RoboDK station: PRBE_Tache_Bras.rdk

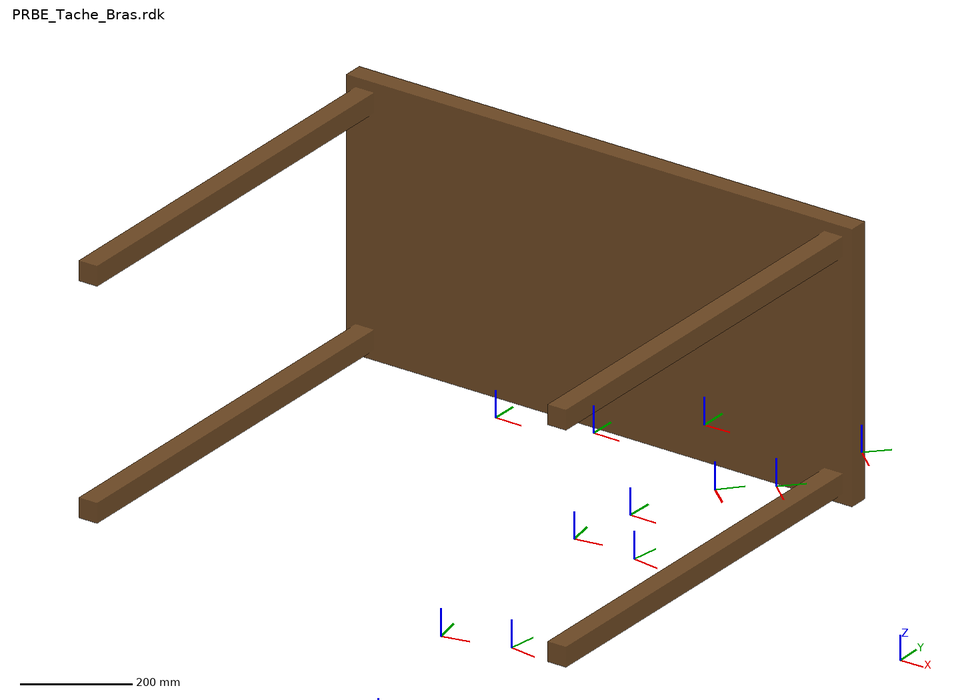
[picture v0: the station drawn from its stored meshes, robots at their saved joint values, targets as dots, program paths as lines]
Station PRBE_Tache_Bras (saved by RoboDK 6.0.4). Poses are relative to the parent item; angles as X-Y-Z fixed-axis rotations.
  - object Manikin_1 at (0, 0, 0) mm, geometry from Manikin_1.STEP
  - frame Human_Base at (0, 958, 0) mm
    - frame hipL_abduction at (63.26, -78.51, -37.42) mm, rotated rx 0 ry 0 rz -7.94 deg
      - frame hipL_flexion at (0, 0, 0) mm
        - frame hipL_rotation at (0, 0, 0) mm
          - frame kneeL_flexion at (67.44, -393.44, -12.97) mm
            - frame ankleL_flexion at (42.46, -394.54, 0) mm, rotated rx 0 ry 0 rz 7.94 deg
              - item type 7 Manikin_1-pied_g
            - item type 7 Manikin_1-tibia_g
          - item type 7 Manikin_1-cuisse_g
    - frame shoulderL_abduction at (206.4, 423.68, 12.96) mm, rotated rx 0 ry 0 rz -42 deg
      - frame shoulderL_flexion at (0, 0, 0) mm
        - frame shoulderL_rotation at (0, 0, 0) mm
          - frame elbowL_flexion at (155.8, -191.9, 27.9) mm
            - frame wristL_flexion at (148.7, -146.81, 80.89) mm
              - frame wristL_deviation at (0, 0, 0) mm
                - item type 7 Manikin_1-main_g
            - item type 7 Manikin_1-avant_bras_g
          - item type 7 Manikin_1-bras_g
    - frame hipR_abduction at (-70.11, -75.34, -37.06) mm, rotated rx 0 ry 0 rz 10.84 deg
      - frame hipR_flexion at (0, 0, 0) mm
        - frame hipR_rotation at (0, 0, 0) mm
          - frame kneeR_flexion at (-86.5, -385.51, -37.91) mm
            - frame ankleR_flexion at (-60.5, -382.31, -26.03) mm, rotated rx 0 ry 0 rz -10.84 deg
              - item type 7 Manikin_1-pied_d_1
              - item type 7 Manikin_1-pied_d_2
            - item type 7 Manikin_1-tibia_d_1
            - item type 7 Manikin_1-tibia_d_2
          - item type 7 Manikin_1-cuisse_d
    - frame shoulderR_abduction at (-133.98, 420.49, -26.02) mm
      - frame shoulderR_flexion at (0, 0, 0) mm
        - frame shoulderR_rotation at (0, 0, 0) mm
          - frame elbowR_flexion at (-80.76, -228.86, 52.14) mm
            - frame wristR_flexion at (-76.34, -195.54, 87.27) mm
              - frame wristR_deviation at (0, 0, 0) mm
                - item type 7 Manikin_1-main_d
            - item type 7 Manikin_1-avant_bras_d
          - item type 7 Manikin_1-bras_d
    - item type 7 Manikin_1-tete
    - item type 7 Manikin_1-bassin
    - item type 7 Manikin_1-torso
  - Python program Marche_Militaire (listed below)
  - Python program Marche_Avant (listed below)
  - Python program Marche_Trajectoire (listed below)
  - Python program fix_reattache_segments (listed below)
  - Python program Position_0 (listed below)
  - object Table at (0, 900, 485) mm, size 1100 x 900 x 550 mm
  - object Trajectoire_Marche at (0, 0, 0) mm
  - Python program Tache_Bras (listed below)
  - object Piece at (80, 940, 300) mm, size 80 x 80 x 80 mm

--- Python program Marche_Militaire ---
# -*- coding: utf-8 -*-
"""
Marche_Militaire.py — L'operateur marque le pas (marche militaire sur place).

A LANCER DANS ROBODK (clic droit > Run) depuis la station avec le rig 22 DDL,
operateur en pose NEUTRE (le script capture le repos au demarrage).

Principe de la marche militaire :
  - genoux qui montent haut, alternes
  - bras RAIDES (coude quasi tendu) qui balancent en OPPOSITION des jambes
  - buste droit (il est fige, parfait pour un militaire)

Regle les amplitudes/vitesse dans la section REGLAGES.
"""
from robolink import Robolink
from robodk.robomath import rotx, roty, rotz
import math
import time

RDK = Robolink()

# ---- Les 22 DDL : nom -> (axe, limite_basse_deg, limite_haute_deg) ----
DDL = {
    # JAMBE DROITE (5)
    "hipR_abduction": ("z", -45, 30),   "hipR_flexion": ("x", -120, 15),  "hipR_rotation": ("y", -45, 45),
    "kneeR_flexion":  ("x", 0, 135),    "ankleR_flexion": ("x", -30, 50),
    # JAMBE GAUCHE (5)
    "hipL_abduction": ("z", -30, 45),   "hipL_flexion": ("x", -120, 15),  "hipL_rotation": ("y", -45, 45),
    "kneeL_flexion":  ("x", 0, 135),    "ankleL_flexion": ("x", -30, 50),
    # BRAS DROIT (6)
    "shoulderR_abduction": ("z", -135, 90), "shoulderR_flexion": ("x", -90, 90), "shoulderR_rotation": ("y", -45, 180),
    "elbowR_flexion": ("x", 0, 145),
    "wristR_flexion": ("x", -50, 60),   "wristR_deviation": ("z", -30, 20),
    # BRAS GAUCHE (6)
    "shoulderL_abduction": ("z", -90, 135), "shoulderL_flexion": ("x", -90, 90), "shoulderL_rotation": ("y", -45, 180),
    "elbowL_flexion": ("x", 0, 145),
    "wristL_flexion": ("x", -50, 60),   "wristL_deviation": ("z", -30, 20),
}

ROT = {"x": rotx, "y": roty, "z": rotz}
F = {nom: RDK.Item(nom) for nom in DDL}            # les reperes
REST = {nom: F[nom].Pose() for nom in DDL}         # pose neutre (capturee au demarrage)


def bouge(nom, deg):
    """Tourne un DDL de `deg` degres depuis le repos (borne aux limites)."""
    axe, lo, hi = DDL[nom]
    deg = max(lo, min(hi, deg))
    F[nom].setPose(REST[nom] * ROT[axe](math.radians(deg)))


def neutre():
    """Remet tout l'operateur droit."""
    for nom in DDL:
        F[nom].setPose(REST[nom])


# =======================================================================
# REGLAGES de la marche militaire
# =======================================================================
HANCHE = 55      # levee de cuisse (deg) — genou haut
GENOU = 65       # pliage du genou quand la jambe monte (deg)
CHEVILLE = 15    # pointe de pied quand la jambe est levee (deg)
BRAS_AV = -45    # bras vers l'AVANT (deg, negatif = devant)
BRAS_ARR = 20    # bras vers l'ARRIERE (deg)
COUDE = 8        # coude quasi tendu = bras raide militaire
NB_PAS = 8       # nombre de pas au total
IMAGES_PAR_PAS = 12   # fluidite (images par pas)
DT = 0.04        # pause entre images (s) — plus petit = plus rapide


def pose_marche(ph):
    """Pose complete de la marche pour une phase `ph` (radians).
       Jambe droite levee sur [0, pi], jambe gauche sur [pi, 2pi]."""
    s = math.sin(ph)
    lift_d = max(0.0, s)     # jambe droite qui monte
    lift_g = max(0.0, -s)    # jambe gauche qui monte

    # jambes : genou haut + pointe de pied
    bouge("hipR_flexion", -HANCHE * lift_d)
    bouge("kneeR_flexion", GENOU * lift_d)
    bouge("ankleR_flexion", CHEVILLE * lift_d)
    bouge("hipL_flexion", -HANCHE * lift_g)
    bouge("kneeL_flexion", GENOU * lift_g)
    bouge("ankleL_flexion", CHEVILLE * lift_g)

    # bras raides, en opposition : bras droit devant quand jambe gauche monte
    u_d = (1.0 - s) / 2.0    # 0 = bras D derriere, 1 = bras D devant
    u_g = (1.0 + s) / 2.0
    bouge("shoulderR_flexion", BRAS_ARR + (BRAS_AV - BRAS_ARR) * u_d)
    bouge("shoulderL_flexion", BRAS_ARR + (BRAS_AV - BRAS_ARR) * u_g)
    bouge("elbowR_flexion", COUDE)
    bouge("elbowL_flexion", COUDE)


def marche(nb_pas=NB_PAS, images_par_pas=IMAGES_PAR_PAS, dt=DT):
    """Anime la marche militaire sur place."""
    for i in range(nb_pas * images_par_pas + 1):
        ph = math.pi * i / images_par_pas      # 1 pas = une demi-periode
        RDK.Render(False)
        pose_marche(ph)
        RDK.Render(True)
        time.sleep(dt)
    neutre()
    RDK.Render(True)


if __name__ == "__main__":
    print("Marche militaire : {} pas...".format(NB_PAS))
    marche()
    print("Repos !")

--- Python program Marche_Avant ---
# -*- coding: utf-8 -*-
"""
Marche_Avant.py — L'operateur marche TOUT DROIT devant lui (marche naturelle).

A LANCER DANS ROBODK (clic droit > Run) depuis la station avec le rig 22 DDL,
operateur au repos / garde-a-vous (le script capture le repos au demarrage).

Principe :
  - hanches qui balancent avant/arriere, genou qui se plie pendant le balance
  - bras souples en opposition des jambes (coude legerement plie)
  - le CORPS AVANCE a la vitesse des pas (longueur de pas calculee depuis
    l'amplitude de hanche) -> pas de glisse visible
  - il marche vers SON regard (+Z monde). A la fin, il REVIENT au centre
    (position d'origine de Human_Base).

Regle les amplitudes/vitesse dans la section REGLAGES.
"""
from robolink import Robolink
from robodk.robomath import rotx, roty, rotz, transl
import math
import time

RDK = Robolink()

# ---- Les 22 DDL : nom -> (axe, limite_basse_deg, limite_haute_deg) ----
DDL = {
    # JAMBE DROITE (5)
    "hipR_abduction": ("z", -45, 30),   "hipR_flexion": ("x", -120, 15),  "hipR_rotation": ("y", -45, 45),
    "kneeR_flexion":  ("x", 0, 135),    "ankleR_flexion": ("x", -30, 50),
    # JAMBE GAUCHE (5)
    "hipL_abduction": ("z", -30, 45),   "hipL_flexion": ("x", -120, 15),  "hipL_rotation": ("y", -45, 45),
    "kneeL_flexion":  ("x", 0, 135),    "ankleL_flexion": ("x", -30, 50),
    # BRAS DROIT (6)
    "shoulderR_abduction": ("z", -135, 90), "shoulderR_flexion": ("x", -90, 90), "shoulderR_rotation": ("y", -45, 180),
    "elbowR_flexion": ("x", 0, 145),
    "wristR_flexion": ("x", -50, 60),   "wristR_deviation": ("z", -30, 20),
    # BRAS GAUCHE (6)
    "shoulderL_abduction": ("z", -90, 135), "shoulderL_flexion": ("x", -90, 90), "shoulderL_rotation": ("y", -45, 180),
    "elbowL_flexion": ("x", 0, 145),
    "wristL_flexion": ("x", -50, 60),   "wristL_deviation": ("z", -30, 20),
}

ROT = {"x": rotx, "y": roty, "z": rotz}
F = {nom: RDK.Item(nom) for nom in DDL}            # les reperes
REST = {nom: F[nom].Pose() for nom in DDL}         # pose de repos (capturee au demarrage)
BASE = RDK.Item("Human_Base")
BASE_REST = BASE.Pose()                            # position de depart du corps
HOME = transl(0, 958, 0)                           # position d'origine (au centre, 1er repere)


def bouge(nom, deg):
    """Tourne un DDL de `deg` degres depuis le repos (borne aux limites)."""
    axe, lo, hi = DDL[nom]
    deg = max(lo, min(hi, deg))
    F[nom].setPose(REST[nom] * ROT[axe](math.radians(deg)))


def neutre():
    """Remet les articulations au repos (le corps reste ou il est)."""
    for nom in DDL:
        F[nom].setPose(REST[nom])


# =======================================================================
# REGLAGES de la marche
# =======================================================================
HANCHE_AV = 30    # jambe vers l'avant (deg)
HANCHE_ARR = 12   # jambe vers l'arriere (deg)
GENOU = 50        # pliage du genou pendant le balance (deg)
CHEVILLE = 8      # pointe de pied relevee pendant le balance (deg)
BRAS_AV = 25      # bras vers l'avant (deg)
BRAS_ARR = 15     # bras vers l'arriere (deg)
COUDE = 20        # coude legerement plie (marche naturelle)
NB_PAS = 8        # nombre de pas
IMAGES_PAR_PAS = 14   # fluidite
DT = 0.04         # pause entre images (s)

LONGUEUR_JAMBE = 790.0   # hanche -> cheville (mm, mesure sur le modele)
SENS = +1                # +1 = devant lui (+Z monde). Mets -1 pour marche arriere.

# longueur d'un pas deduite du balancement de hanche (pour avancer sans glisser)
LONGUEUR_PAS = LONGUEUR_JAMBE * (math.sin(math.radians(HANCHE_AV)) + math.sin(math.radians(HANCHE_ARR)))


def pose_pas(ph):
    """Pose de marche pour une phase `ph` (radians). Jambe droite devant sur [0, pi]."""
    s = math.sin(ph)
    # hanches : avant = negatif (amplitude asymetrique avant/arriere)
    a = (HANCHE_AV + HANCHE_ARR) / 2.0
    c = (HANCHE_AV - HANCHE_ARR) / 2.0
    bouge("hipR_flexion", -(a * s + c))
    bouge("hipL_flexion", -(a * -s + c))
    # genou plie pendant le balance (jambe qui revient vers l'avant)
    bouge("kneeR_flexion", GENOU * max(0.0, math.cos(ph)))
    bouge("kneeL_flexion", GENOU * max(0.0, -math.cos(ph)))
    # pointe de pied relevee pendant le balance (pour ne pas racler le sol)
    bouge("ankleR_flexion", -CHEVILLE * max(0.0, math.cos(ph)))
    bouge("ankleL_flexion", -CHEVILLE * max(0.0, -math.cos(ph)))
    # bras en opposition, coude souple
    sa = (BRAS_AV + BRAS_ARR) / 2.0
    sc = (BRAS_ARR - BRAS_AV) / 2.0
    bouge("shoulderR_flexion", sa * s + sc)
    bouge("shoulderL_flexion", -sa * s + sc)
    bouge("elbowR_flexion", COUDE)
    bouge("elbowL_flexion", COUDE)


def avance(dist):
    """Place le corps a `dist` mm devant sa position de depart."""
    BASE.setPose(BASE_REST * transl(0, 0, SENS * dist))


def marche(nb_pas=NB_PAS, images_par_pas=IMAGES_PAR_PAS, dt=DT):
    """Anime la marche en avant, puis remet l'operateur au centre (HOME)."""
    for i in range(nb_pas * images_par_pas + 1):
        ph = math.pi * i / images_par_pas      # 1 pas = une demi-periode
        RDK.Render(False)
        pose_pas(ph)
        avance(LONGUEUR_PAS * ph / math.pi)
        RDK.Render(True)
        time.sleep(dt)
    # fin : repos + retour a la position initiale, au centre
    RDK.Render(False)
    neutre()
    BASE.setPose(HOME)
    RDK.Render(True)


if __name__ == "__main__":
    d_tot = LONGUEUR_PAS * NB_PAS / 1000.0
    print("Marche avant : {} pas (~{:.1f} m)...".format(NB_PAS, d_tot))
    marche()
    print("Arrive !")

--- Python program Marche_Trajectoire ---
# -*- coding: utf-8 -*-
"""
Marche_Trajectoire.py — L'operateur marche le long d'une TRAJECTOIRE EXTERNE
(non lineaire), definie par des waypoints dans un fichier JSON.

A LANCER DANS ROBODK (clic droit > Run) depuis la station avec le rig 22 DDL,
operateur au repos / garde-a-vous (le script capture le repos au demarrage).

Principe (demande reunion du 04/06) :
  - la trajectoire est DEFINIE EN EXTERNE : trajectoires\\trajectoire_S.json
    (liste de points [x, z] au sol, en mm) -> modifiable sans toucher au code
  - les waypoints sont lisses par une spline Catmull-Rom -> courbe douce
  - le corps SUIT la courbe par abscisse curviligne : position sur la courbe
    + orientation vers la tangente (il regarde toujours ou il va)
  - meme cycle de marche et meme anti-glisse que Marche_Avant : le corps
    avance a la vitesse des pas (longueur de pas deduite du balancement
    de hanche), donc pas de patinage le long de la courbe
  - la trajectoire est tracee au sol dans la station (courbe bleue)

Usage terminal (RoboDK ouvert) :
    python Marche_Trajectoire.py [chemin\\trajectoire.json] [--reste]
    --reste : ne pas revenir au centre a la fin (rester au bout du chemin)
"""
from robolink import Robolink
from robodk.robomath import rotx, roty, rotz, transl
import bisect
import json
import math
import sys
import time

RDK = Robolink()

# ---- Les 22 DDL : nom -> (axe, limite_basse_deg, limite_haute_deg) ----
DDL = {
    # JAMBE DROITE (5)
    "hipR_abduction": ("z", -45, 30),   "hipR_flexion": ("x", -120, 15),  "hipR_rotation": ("y", -45, 45),
    "kneeR_flexion":  ("x", 0, 135),    "ankleR_flexion": ("x", -30, 50),
    # JAMBE GAUCHE (5)
    "hipL_abduction": ("z", -30, 45),   "hipL_flexion": ("x", -120, 15),  "hipL_rotation": ("y", -45, 45),
    "kneeL_flexion":  ("x", 0, 135),    "ankleL_flexion": ("x", -30, 50),
    # BRAS DROIT (6)
    "shoulderR_abduction": ("z", -135, 90), "shoulderR_flexion": ("x", -90, 90), "shoulderR_rotation": ("y", -45, 180),
    "elbowR_flexion": ("x", 0, 145),
    "wristR_flexion": ("x", -50, 60),   "wristR_deviation": ("z", -30, 20),
    # BRAS GAUCHE (6)
    "shoulderL_abduction": ("z", -90, 135), "shoulderL_flexion": ("x", -90, 90), "shoulderL_rotation": ("y", -45, 180),
    "elbowL_flexion": ("x", 0, 145),
    "wristL_flexion": ("x", -50, 60),   "wristL_deviation": ("z", -30, 20),
}

ROT = {"x": rotx, "y": roty, "z": rotz}
F = {nom: RDK.Item(nom) for nom in DDL}            # les reperes
REST = {nom: F[nom].Pose() for nom in DDL}         # pose de repos (capturee au demarrage)
BASE = RDK.Item("Human_Base")
HOME = transl(0, 958, 0)                           # position d'origine (au centre)
Y0 = BASE.Pose().Pos()[1]                          # hauteur du bassin (958 mm)


def bouge(nom, deg):
    """Tourne un DDL de `deg` degres depuis le repos (borne aux limites)."""
    axe, lo, hi = DDL[nom]
    deg = max(lo, min(hi, deg))
    F[nom].setPose(REST[nom] * ROT[axe](math.radians(deg)))


def neutre():
    """Remet les articulations au repos (le corps reste ou il est)."""
    for nom in DDL:
        F[nom].setPose(REST[nom])


# =======================================================================
# REGLAGES
# =======================================================================
TRAJET_DEFAUT = r"D:\PRBE_Homme_Robot\PRBE-Homme-Robot\trajectoires\trajectoire_S.json"
HANCHE_AV = 30    # jambe vers l'avant (deg)
HANCHE_ARR = 12   # jambe vers l'arriere (deg)
GENOU = 50        # pliage du genou pendant le balance (deg)
CHEVILLE = 8      # pointe de pied relevee pendant le balance (deg)
BRAS_AV = 25      # bras vers l'avant (deg)
BRAS_ARR = 15     # bras vers l'arriere (deg)
COUDE = 20        # coude legerement plie
IMAGES_PAR_PAS = 14   # fluidite
DT = 0.04         # pause entre images (s)
TRACER = True     # dessiner la trajectoire au sol dans la station

LONGUEUR_JAMBE = 790.0   # hanche -> cheville (mm)
LONGUEUR_PAS = LONGUEUR_JAMBE * (math.sin(math.radians(HANCHE_AV)) + math.sin(math.radians(HANCHE_ARR)))


# =======================================================================
# Trajectoire : JSON -> spline Catmull-Rom -> abscisse curviligne
# =======================================================================
def charge_waypoints(chemin):
    with open(chemin, encoding="utf-8") as f:
        data = json.load(f)
    pts = [tuple(map(float, p)) for p in data["points_xz_mm"]]
    if len(pts) < 2:
        raise SystemExit("ERREUR : il faut au moins 2 waypoints.")
    return data.get("nom", "(sans nom)"), pts


def _cr(p0, p1, p2, p3, t):
    """Point de Catmull-Rom (uniforme) entre p1 et p2, t dans [0,1]."""
    t2, t3 = t * t, t * t * t
    return tuple(0.5 * (2 * p1[k] + (-p0[k] + p2[k]) * t
                        + (2 * p0[k] - 5 * p1[k] + 4 * p2[k] - p3[k]) * t2
                        + (-p0[k] + 3 * p1[k] - 3 * p2[k] + p3[k]) * t3)
                 for k in range(2))


def lisse(waypoints, par_segment=24):
    """Spline Catmull-Rom a travers les waypoints -> polyligne dense."""
    P = [waypoints[0]] + list(waypoints) + [waypoints[-1]]
    dense = []
    for i in range(len(waypoints) - 1):
        for j in range(par_segment):
            dense.append(_cr(P[i], P[i + 1], P[i + 2], P[i + 3], j / par_segment))
    dense.append(waypoints[-1])
    return dense


def abscisses(dense):
    """Longueurs cumulees le long de la polyligne."""
    S = [0.0]
    for a, b in zip(dense, dense[1:]):
        S.append(S[-1] + math.hypot(b[0] - a[0], b[1] - a[1]))
    return S


def point_et_tangente(dense, S, s):
    """Position (x,z) + tangente unitaire (tx,tz) a l'abscisse s (mm)."""
    s = max(0.0, min(S[-1], s))
    i = min(max(bisect.bisect_left(S, s), 1), len(S) - 1)
    seg = S[i] - S[i - 1] or 1e-9
    u = (s - S[i - 1]) / seg
    a, b = dense[i - 1], dense[i]
    x = a[0] + u * (b[0] - a[0])
    z = a[1] + u * (b[1] - a[1])
    tx, tz = b[0] - a[0], b[1] - a[1]
    n = math.hypot(tx, tz) or 1e-9
    return (x, z), (tx / n, tz / n)


def tracer_trajectoire(dense):
    """Dessine la courbe au sol dans la station (best effort)."""
    try:
        vieux = RDK.Item("Trajectoire_Marche")
        if vieux.Valid() and vieux.Name() == "Trajectoire_Marche":
            vieux.Delete()
        courbe = RDK.AddCurve([[p[0], 10.0, p[1]] for p in dense])
        if courbe.Valid():
            courbe.setName("Trajectoire_Marche")
            courbe.setColorCurve([0.1, 0.3, 0.9, 1])
    except Exception as e:  # noqa: BLE001
        print("(trace de la trajectoire ignoree : {})".format(e))


# =======================================================================
# Cycle de marche (identique a Marche_Avant)
# =======================================================================
def pose_pas(ph):
    """Pose de marche pour une phase `ph` (radians). Jambe droite devant sur [0, pi]."""
    s = math.sin(ph)
    a = (HANCHE_AV + HANCHE_ARR) / 2.0
    c = (HANCHE_AV - HANCHE_ARR) / 2.0
    bouge("hipR_flexion", -(a * s + c))
    bouge("hipL_flexion", -(a * -s + c))
    bouge("kneeR_flexion", GENOU * max(0.0, math.cos(ph)))
    bouge("kneeL_flexion", GENOU * max(0.0, -math.cos(ph)))
    bouge("ankleR_flexion", -CHEVILLE * max(0.0, math.cos(ph)))
    bouge("ankleL_flexion", -CHEVILLE * max(0.0, -math.cos(ph)))
    sa = (BRAS_AV + BRAS_ARR) / 2.0
    sc = (BRAS_ARR - BRAS_AV) / 2.0
    bouge("shoulderR_flexion", sa * s + sc)
    bouge("shoulderL_flexion", -sa * s + sc)
    bouge("elbowR_flexion", COUDE)
    bouge("elbowL_flexion", COUDE)


def place_corps(dense, S, s):
    """Place le corps a l'abscisse s : position sur la courbe + regard tangent."""
    (x, z), (tx, tz) = point_et_tangente(dense, S, s)
    theta = math.atan2(tx, tz)          # le mannequin regarde vers +Z local
    BASE.setPose(transl(x, Y0, z) * roty(theta))


def marche_trajectoire(dense, S, retour_centre=True):
    """Anime la marche le long de la courbe, du debut a la fin."""
    L = S[-1]
    nb_images = int(math.ceil(L / LONGUEUR_PAS * IMAGES_PAR_PAS))
    for i in range(nb_images + 1):
        ph = math.pi * i / IMAGES_PAR_PAS          # 1 pas = une demi-periode
        s = min(L, LONGUEUR_PAS * ph / math.pi)    # anti-glisse : s = vitesse des pas
        RDK.Render(False)
        pose_pas(ph)
        place_corps(dense, S, s)
        RDK.Render(True)
        time.sleep(DT)
    # fin : repos (oriente comme a l'arrivee)
    RDK.Render(False)
    neutre()
    if retour_centre:
        BASE.setPose(HOME)
    RDK.Render(True)


if __name__ == "__main__":
    args = [a for a in sys.argv[1:] if a != "--reste"]
    reste = "--reste" in sys.argv[1:]
    chemin = args[0] if args else TRAJET_DEFAUT

    nom, waypoints = charge_waypoints(chemin)
    dense = lisse(waypoints)
    S = abscisses(dense)
    if TRACER:
        tracer_trajectoire(dense)
    print("Trajectoire '{}' : {} waypoints, {:.1f} m, ~{} pas".format(
        nom, len(waypoints), S[-1] / 1000.0, int(round(S[-1] / LONGUEUR_PAS))))
    marche_trajectoire(dense, S, retour_centre=not reste)
    p = BASE.Pose().Pos()
    print("Arrive ! Position finale Human_Base : x={:.0f} y={:.0f} z={:.0f} (retour_centre={})".format(
        p[0], p[1], p[2], not reste))

--- Python program fix_reattache_segments ---
# -*- coding: utf-8 -*-
"""
fix_reattache_segments.py — Repare le mannequin eclate a la reouverture du
.rdk SANS rebuild (quelques secondes), en re-jouant le re-basage geometrique
perdu a la sauvegarde.

Cause (diagnostic du 10/06) : pour les sous-solides type 7 (courbes issues
du Split), le .rdk sauve les points BRUTS d'origine — la compensation posee
par setParentStatic au moment du rig n'est PAS persistee. A l'ouverture,
RoboDK applique la transformation du frame parent sur ces points bruts
-> double transformation -> mannequin eclate. Les frames, vrais items a
pose persistee, restent corrects.

Remede, segment par segment :
  1) memoriser la pose relative de chaque frame, puis remettre chaque
     frame en etat de CONSTRUCTION (translation seule, rotation identite —
     l'etat dans lequel le rig d'origine a pose ses compensations)
  2) setParent(station)      — detache en KEEP-RELATIVE : la compensation
     (identite au chargement) ne change pas -> le segment retombe sur ses
     points bruts = position d'import, mannequin recompose
     setParentStatic(frame)  — re-attache en preservant l'absolu : la
     compensation F_build^-1 est re-posee, exactement comme au rig
  3) restaurer les poses memorisees (garde-a-vous, jambes resserrees) :
     la geometrie suit les frames

!! NE PAS envelopper dans RDK.Render(False) : le re-basage des type 7
echoue silencieusement sans rendu actif (constate le 10/06 — deux
tentatives identiques en Render(False) = aucun effet, la meme sequence
render actif fonctionne).

A relancer A CHAQUE OUVERTURE du .rdk (la sauvegarde re-perd le re-basage).
Filet de securite si etat incoherent : scripts/rebuild_operateur.py (~30 s).

!! PAS IDEMPOTENT : sur une station SAINE (fraichement rebuildee ou deja
reparee), le re-basage s'appliquerait une fois de trop et eclaterait le
mannequin. Une garde detecte l'etat via un segment du tronc et refuse de
tourner si la station est saine (--force pour outrepasser).

Usage (RoboDK ouvert, station chargee) :
    python fix_reattache_segments.py [--skip nom1,nom2] [--force]
    --skip  : segments a ne pas toucher (ex. deja repares a la main)
    --force : sauter la garde de detection
"""
import math
import sys
import time
from pathlib import Path
sys.path.insert(0, str(Path(__file__).resolve().parent))
from robolink import Robolink, ITEM_TYPE_FRAME
from robodk.robomath import transl

# ancres d'import des segments du tronc (cf. build_human_robodk.ANCHORS),
# en dur pour que le script reste autonome une fois embarque dans la station
TRONC = {"tete": (20, 1584, 30), "torso": (15, 1260, 0), "bassin": (0, 958, 0)}

skip = set()
if "--skip" in sys.argv:
    skip = set(sys.argv[sys.argv.index("--skip") + 1].split(","))

t0 = time.time()
RDK = Robolink()
station = RDK.ActiveStation()
print("Station :", station.Name())


def _d(a, b):
    return math.sqrt(sum((x - y) ** 2 for x, y in zip(a, b)))


def garde_station_cassee():
    """True si le mannequin est eclate (double transformation detectee)."""
    for it in RDK.ItemList():
        if it.Type() != 7:
            continue
        part = it.Name().split("-", 1)[-1]
        if part not in TRONC:
            continue
        bb = it.setParam("BoundingBox")
        c = [(bb["min"][i] + bb["max"][i]) / 2.0 for i in range(3)]
        a = TRONC[part]
        F = it.Parent().PoseAbs().rows
        fa = [sum(F[i][j] * a[j] for j in range(3)) + F[i][3] for i in range(3)]
        d_sain, d_casse = _d(c, a), _d(c, fa)
        etat = "CASSEE (double transformation)" if d_casse < d_sain else "saine"
        print(f"Garde ({part}) : d_sain={d_sain:.0f} mm, d_casse={d_casse:.0f} mm -> station {etat}")
        return d_casse < d_sain
    sys.exit("Garde impossible : aucun segment du tronc (tete/torso/bassin) trouve.")


if "--force" not in sys.argv and not garde_station_cassee():
    sys.exit("Rien a faire — relancer avec --force pour outrepasser la garde.")

frames = RDK.ItemList(ITEM_TYPE_FRAME)
solids = [it for it in RDK.ItemList() if it.Type() == 7]
if not solids:
    sys.exit("Rien a reparer : aucun sous-solide type 7 dans la station.")
parent_of = {}
for s in solids:
    nm = s.Name()
    if nm in skip or nm.split("-", 1)[-1] in skip:
        print(f"  (skip : {nm})")
        continue
    p = s.Parent()
    if p.Type() == 3:
        parent_of[s] = p
    else:
        print(f"  (ignore : {nm} n'est pas sous un frame)")
print(f"{len(frames)} frames, {len(parent_of)} segments a re-attacher")

# 1) frames -> etat de construction (translation seule)
saved = []
for fr in frames:
    pose = fr.Pose()
    saved.append((fr, pose))
    r = pose.rows
    fr.setPose(transl(r[0][3], r[1][3], r[2][3]))

# 2) re-basage : detacher en keep-relative, re-attacher en statique
for s, fr in parent_of.items():
    s.setParent(station)
    s.setParentStatic(fr)
    print(f"  re-attache : {s.Name():26s} -> {fr.Name()}")

# 3) restaurer les poses (garde-a-vous, jambes resserrees, ...)
for fr, pose in saved:
    fr.setPose(pose)

print(f"OK — {len(parent_of)} segments re-attaches en {time.time() - t0:.1f} s")

--- Python program Position_0 ---
# -*- coding: utf-8 -*-
"""
Position_0.py — Remet le mannequin au GARDE-A-VOUS exact (position zero).

A lancer quand on veut repartir d'un etat propre : apres une animation
interrompue, un script qui a laisse le bras en l'air, ou des residus
accumules (chaque animation se termine a quelques degres pres ; les petits
ecarts s'additionnent au fil des runs).

Reconstruit le zero du rig (cf. rig_active_station.py, section 8) :
  - les 22 DDL -> rotation IDENTITE (la translation du repere ne bouge
    jamais, on la conserve telle quelle) ;
  - epaule du cote X+ (= gauche) : rotz(-42 deg) pour plaquer le bras que
    la pose STEP d'origine ecarte du corps ;
  - jambes resserrees : cheville ramenee a l'aplomb de la hanche (angle
    recalcule depuis les positions des reperes, pied contre-tourne).

Ne touche ni la Table, ni la Piece, ni la camera.
    C:\\RoboDK\\Python-Embedded\\python.exe scripts\\Position_0.py
"""
import math
import sys
from robolink import Robolink, ITEM_TYPE_FRAME
from robodk.robomath import Mat, rotz

RDK = Robolink()
print("Station :", RDK.ActiveStation().Name())

DOF = [
    "shoulderL_abduction", "shoulderL_flexion", "shoulderL_rotation",
    "elbowL_flexion", "wristL_flexion", "wristL_deviation",
    "shoulderR_abduction", "shoulderR_flexion", "shoulderR_rotation",
    "elbowR_flexion", "wristR_flexion", "wristR_deviation",
    "hipL_abduction", "hipL_flexion", "hipL_rotation", "kneeL_flexion",
    "ankleL_flexion",
    "hipR_abduction", "hipR_flexion", "hipR_rotation", "kneeR_flexion",
    "ankleR_flexion",
]

F = {}
for nm in DOF:
    fr = RDK.Item(nm, ITEM_TYPE_FRAME)
    if not fr.Valid():
        sys.exit(f"ERREUR : repere {nm} introuvable — rig 22 DDL absent ?")
    F[nm] = fr


def zero(fr):
    """Rotation identite, translation conservee."""
    p = fr.Pose()
    fr.setPose(Mat([[1, 0, 0, p[0, 3]], [0, 1, 0, p[1, 3]],
                    [0, 0, 1, p[2, 3]], [0, 0, 0, 1]]))


# 1) tout a zero (les positions absolues redeviennent celles de la pose STEP)
for nm in DOF:
    zero(F[nm])

# 2) bras gauche (cote X+) plaque le long du corps
F["shoulderL_abduction"].setPose(
    F["shoulderL_abduction"].Pose() * rotz(math.radians(-42.0)))

# 3) jambes resserrees : meme calcul que le rig (cheville a l'aplomb de la
#    hanche), possible car a l'etape 1 les reperes sont aux positions STEP
for u in ("R", "L"):
    hp = F[f"hip{u}_abduction"].PoseAbs()
    ap = F[f"ankle{u}_flexion"].PoseAbs()
    ang = math.atan2(ap[0, 3] - hp[0, 3], hp[1, 3] - ap[1, 3])
    F[f"hip{u}_abduction"].setPose(F[f"hip{u}_abduction"].Pose() * rotz(-ang))
    F[f"ankle{u}_flexion"].setPose(F[f"ankle{u}_flexion"].Pose() * rotz(ang))
    print(f"  jambes resserrees ({u}) : {math.degrees(ang):+.1f} deg")

RDK.Render(True)
print("Position 0 : mannequin au garde-a-vous.")

--- Python program Tache_Bras ---
# -*- coding: utf-8 -*-
"""
Tache_Bras.py — v3 (refonte complete, 11/06) : pick & place d'une piece
cubique sur une table, bras gauche 6 DDL, corps fixe.

Scenario :
  Le mannequin est debout devant une table. Une piece cubique est posee
  pres du BORD AVANT de la table, a sa GAUCHE. Il la saisit de la main
  gauche, la deplace vers la DROITE et la repose sur la meme table.

REGLES v3 (retours Niko 11/06, "reprendre a zero") :

  1. LE COUDE PART EN ARRIERE, JAMAIS EN AVANT. La position du coude ne
     depend que de l'epaule ; sur ce rig la flexion d'epaule POSITIVE le
     tire en arriere (sonde _probe_coude : flexion +10 => coude Z 41->7).
     La flexion est donc BORNEE a [-8, +25] pour TOUT le scenario : le
     bras ne bascule jamais vers l'avant, la main avance par le pli du
     coude. Consequence geometrique : la piece doit etre pres du bord
     avant de la table (Z=300 et non 400 — a 400 il FAUT avancer le
     coude, c'est ce qui pourrissait la v2). Verification integree :
     le Z du coude est scanne sur TOUTE la trajectoire precalculee.

  2. MOUVEMENT DYNAMIQUE. La lenteur de la v2 venait de l'IK calculee A
     CHAQUE FRAME pendant l'animation (~400 appels FK par image). La v3
     PRECALCULE toute la trajectoire articulaire (IK seulement sur les
     postures cles, hors animation), puis la JOUE a cadence fixe : zero
     calcul pendant la lecture, vitesses articulaires ~80-140 deg/s
     (rythme humain), profil doux (smoothstep) par phase, micro-pauses
     saisie/depose.

A LANCER : RoboDK ouvert, station avec le rig 22 DDL.
    C:\\RoboDK\\Python-Embedded\\python.exe scripts\\Tache_Bras.py
    options : --check (precalcul + verifs seulement, pas d'animation)
              --frames (laisser les reperes visibles)

Convention station : X+ = cote GAUCHE du mannequin, +Z = devant, Y = haut.
"""
import math
import sys
import time
from pathlib import Path
sys.path.insert(0, str(Path(__file__).resolve().parent))
# version embarquee dans la station : __file__ pointe vers un dossier temp,
# il faut le chemin absolu du repo pour trouver Position_0
sys.path.insert(0, r"D:\PRBE_Homme_Robot\PRBE-Homme-Robot\scripts")
from robolink import Robolink, ITEM_TYPE_FRAME
from robodk.robomath import Mat, transl, rotx, roty, rotz, invH

# ---------------- parametres de la scene (mm) ----------------
TABLE_TOP = 900          # hauteur de la surface de la table
TABLE_SX, TABLE_SZ = 1100, 550   # plateau : largeur (X) x profondeur (Z)
TABLE_TH = 40            # epaisseur plateau
TABLE_CZ = 485           # centre du plateau devant le mannequin (Z)
CUBE = 80                # arete de la piece cubique
PICK_X, PICK_Z = 330, 300        # piece au depart : a GAUCHE, pres du bord
PLACE_X, PLACE_Z = 80, 300       # depose : 25 cm vers la DROITE, meme bord
                                 # (bord avant : seule zone atteignable
                                 # avec le coude qui reste en ARRIERE)
GRASP_CLEAR = 35         # centre de la main au-dessus du haut du cube (saisie)
HI = 1030                # hauteur de transit (centre paume) : plafond
                         # atteignable coude en arriere. Cube et doigts a
                         # paume-115 = 915, soit ~15 mm au-dessus du
                         # plateau : la piece GLISSE juste au-dessus de la
                         # table — le geste humain pour 25 cm de deport
                         # (on ne souleve pas a 15 cm), valide au mesh
TRANSIT_Z = 280          # transit legerement RAMENE vers le corps (geste
                         # humain : on porte pres de soi) — et plus
                         # atteignable que Z=300 a cette hauteur
DT = 0.025               # cadence de lecture (s/frame) — la trajectoire est
                         # precalculee, la lecture ne fait QUE appliquer+rendre

# ---------------- bras gauche : DDL, axes, limites (deg) ----------------
ARM = [
    ("shoulderL_abduction", "z", -90, 135),
    ("shoulderL_flexion",   "x", -120, 90),
    ("shoulderL_rotation",  "y", -45, 180),
    ("elbowL_flexion",      "x", -145, 0),    # NEGATIF = plier vers l'AVANT
    ("wristL_flexion",      "x", -50, 60),
    ("wristL_deviation",    "z", -30, 20),
]
ROT = {"x": rotx, "y": roty, "z": rotz}

# Bornes du scenario. LA contrainte v3 est la FLEXION D'EPAULE >= -8 :
# le bras ne bascule jamais en avant => le coude ne part jamais en avant
# (verifie en plus par le scan coude sur la trajectoire complete).
# Vers l'ARRIERE en revanche on autorise large (+38, extension humaine
# ~45-60) : c'est ce qui donne la hauteur de transit coude recule.
LIM_SCEN = [(-45, 25), (-8, 38), (-45, 60), (-130, 0), (-40, 55), (-25, 20)]

# ORIENTATION DE LA MAIN : le bras n'a pas de pronation d'avant-bras, on
# garde la main dans son orientation de repos (verticale, doigts vers le
# bas) = identite du repere poignet. Stricte quand la main PORTE la piece,
# souple a main vide.
R_GRASP = Mat([[1.0, 0.0, 0.0, 0.0],
               [0.0, 1.0, 0.0, 0.0],
               [0.0, 0.0, 1.0, 0.0],
               [0.0, 0.0, 0.0, 1.0]])
WO = 65.0           # poids orientation stricte (mm equivalents par radian)
WO_LIBRE = 22.0     # orientation souple (main vide)
LAM = 5.0           # amortissement DLS

# Posture de confort (tache secondaire de l'IK) : selectionne la branche
# "coude en arriere" — epaule legerement en extension, coude plie.
Q_CONF = [0.0, 12.0, 15.0, -80.0, 0.0, 0.0]
WQ = 1.2

RDK = Robolink()
print("Station :", RDK.ActiveStation().Name())

# Remise a zero AVANT de capturer le repos (sinon les residus d'une
# animation precedente corrompent tout le modele FK).
from Position_0 import remettre_a_zero
remettre_a_zero(RDK, verbose=False)
print("Mannequin remis a zero (garde-a-vous).")


# ---------------- scene : table + piece ----------------

def _box_tris(sx, sy, sz):
    """12 triangles d'un pave centre sur l'origine de l'objet."""
    x, y, z = sx / 2.0, sy / 2.0, sz / 2.0
    v = [(-x, -y, -z), (x, -y, -z), (x, y, -z), (-x, y, -z),
         (-x, -y, z), (x, -y, z), (x, y, z), (-x, y, z)]
    quads = [(0, 1, 2, 3), (4, 7, 6, 5), (0, 4, 5, 1),
             (3, 2, 6, 7), (0, 3, 7, 4), (1, 5, 6, 2)]
    tris = []
    for a, b, c, d in quads:
        tris += [v[a], v[b], v[c], v[a], v[c], v[d]]
    return tris


def _add_box(name, sx, sy, sz, pos, color):
    it = RDK.Item(name)
    if it.Valid() and it.Type() == 5:
        return it
    tris = []
    if name == "Table":
        # plateau (origine objet = centre de la SURFACE du plateau)
        for p in _box_tris(sx, TABLE_TH, sz):
            tris.append((p[0], p[1] - TABLE_TH / 2.0, p[2]))
        # 4 pieds
        for px, pz in ((sx/2-40, sz/2-40), (-(sx/2-40), sz/2-40),
                       (sx/2-40, -(sz/2-40)), (-(sx/2-40), -(sz/2-40))):
            for p in _box_tris(40, TABLE_TOP - TABLE_TH, 40):
                tris.append((p[0] + px, p[1] - TABLE_TH - (TABLE_TOP - TABLE_TH)/2.0, p[2] + pz))
    else:
        tris = _box_tris(sx, sy, sz)
    obj = RDK.AddShape([list(p) for p in tris])
    obj.setName(name)
    obj.setColor(color)
    obj.setPose(transl(*pos))
    return obj


table = _add_box("Table", TABLE_SX, TABLE_TOP, TABLE_SZ,
                 (0, TABLE_TOP, TABLE_CZ), [0.55, 0.38, 0.21, 1])
piece = _add_box("Piece", CUBE, CUBE, CUBE,
                 (PICK_X, TABLE_TOP + CUBE / 2.0, PICK_Z), [0.95, 0.55, 0.10, 1])
print("Scene : Table + Piece en place")

# ---------------- modele FK du bras gauche ----------------
F = {nom: RDK.Item(nom, ITEM_TYPE_FRAME) for nom, *_ in ARM}
for nom, fr in F.items():
    if not fr.Valid():
        sys.exit(f"ERREUR : frame {nom} introuvable — rig 22 DDL absent ?")
REST = {nom: F[nom].Pose() for nom, *_ in ARM}
ROOT = F[ARM[0][0]].Parent().PoseAbs()     # pose absolue du parent de l'epaule

# effecteur : centre de la paume au repos, exprime dans le dernier frame
main = None
for it in RDK.ItemList():
    if it.Type() == 7 and it.Name() == "Manikin_1-main_g":
        main = it
if main is None:
    sys.exit("ERREUR : Manikin_1-main_g introuvable.")
bb = main.setParam("BoundingBox")
hand0 = [(bb["min"][i] + bb["max"][i]) / 2.0 for i in range(3)]
wrist_abs0 = F[ARM[-1][0]].PoseAbs()
E_LOCAL = invH(wrist_abs0) * transl(*hand0)
e = E_LOCAL.rows
E_LOCAL = (e[0][3], e[1][3], e[2][3])
print(f"Effecteur (paume) au repos : ({hand0[0]:.0f}, {hand0[1]:.0f}, {hand0[2]:.0f})")


def fk_pose(q):
    """Pose absolue (Mat 4x4) du repere POIGNET pour les 6 angles q (deg)."""
    P = ROOT
    for (nom, axe, lo, hi), a in zip(ARM, q):
        P = P * REST[nom] * ROT[axe](math.radians(a))
    return P


def fk_coude(q):
    """Position absolue du repere COUDE (ne depend que des 3 DDL epaule)."""
    P = ROOT
    for (nom, axe, lo, hi), a in zip(ARM[:3], q[:3]):
        P = P * REST[nom] * ROT[axe](math.radians(a))
    P = P * REST["elbowL_flexion"]
    r = P.rows
    return [r[0][3], r[1][3], r[2][3]]


def eff_pos(P):
    """Position monde de l'effecteur (centre paume) depuis la pose poignet."""
    r = (P * transl(*E_LOCAL)).rows
    return [r[0][3], r[1][3], r[2][3]]


def cols(M):
    r = M.rows
    return [[r[0][c], r[1][c], r[2][c]] for c in range(3)]


def cross(a, b):
    return [a[1]*b[2]-a[2]*b[1], a[2]*b[0]-a[0]*b[2], a[0]*b[1]-a[1]*b[0]]


def ori_err(Rc, Rd):
    """Erreur d'orientation (vecteur monde, ~rad) menant Rc -> Rd."""
    e = [0.0, 0.0, 0.0]
    for k in range(3):
        c = cross(Rc[k], Rd[k])
        e = [e[i] + c[i] for i in range(3)]
    return [0.5 * v for v in e]


RG = cols(R_GRASP)


def clamp(q):
    return [max(lo, min(hi, a)) for (lo, hi), a in zip(LIM_SCEN, q)]


def _solve6(A, b):
    """Resout A y = b (6x6) par elimination de Gauss avec pivot partiel."""
    n = 6
    M = [row[:] + [b[i]] for i, row in enumerate(A)]
    for c in range(n):
        p = max(range(c, n), key=lambda r: abs(M[r][c]))
        M[c], M[p] = M[p], M[c]
        piv = M[c][c]
        if abs(piv) < 1e-12:
            continue
        for r in range(n):
            if r != c and M[r][c]:
                f = M[r][c] / piv
                M[r] = [M[r][k] - f * M[c][k] for k in range(n + 1)]
    return [M[i][n] / M[i][i] if abs(M[i][i]) > 1e-12 else 0.0 for i in range(n)]


def ik(tpos, q0, tol_p=6.0, tol_o=0.09, iters=240, patience=22, wo=WO):
    """IK 6 DOF position + orientation, DLS amortie, posture secondaire
    Q_CONF (branche coude en arriere). Bornee par LIM_SCEN => la flexion
    d'epaule ne peut JAMAIS depasser +25/-8 : le coude reste en arriere
    par construction. Retourne (q, residu_pos_mm, residu_ori_deg)."""
    q = clamp(list(q0))
    best_q, best_s, stale = q[:], 1e18, 0
    for _ in range(iters):
        P = fk_pose(q)
        p = eff_pos(P)
        Rc = cols(P)
        ep = [tpos[i] - p[i] for i in range(3)]
        eo = ori_err(Rc, RG)
        np_ = math.sqrt(sum(v*v for v in ep))
        no_ = math.sqrt(sum(v*v for v in eo))
        s = np_ + wo * no_
        if s < best_s - 0.05:
            best_s, best_q, stale = s, q[:], 0
        else:
            stale += 1
        if np_ < tol_p and no_ < tol_o:
            return q, np_, math.degrees(no_)
        if stale >= patience:
            break
        x = ep + [wo * v for v in eo]
        # Jacobien 6x6 par differences finies
        J = [[0.0] * 6 for _ in range(6)]
        for j in range(6):
            dq = list(q)
            dq[j] += 0.5
            Pj = fk_pose(dq)
            pj = eff_pos(Pj)
            dphi = ori_err(Rc, cols(Pj))
            for i in range(3):
                J[i][j] = (pj[i] - p[i]) / 0.5
                J[3 + i][j] = wo * dphi[i] / 0.5
        # DLS + tache posturale secondaire (s'estompe pres de la cible)
        wq2 = (WQ * min(1.0, np_ / 60.0)) ** 2
        reg = LAM * LAM + wq2
        JTJ = [[sum(J[k][i] * J[k][r] for k in range(6)) + (reg if i == r else 0)
                for r in range(6)] for i in range(6)]
        b = [sum(J[k][j] * x[k] for k in range(6)) + wq2 * (Q_CONF[j] - q[j])
             for j in range(6)]
        dq = _solve6(JTJ, b)
        # rebroussement si le pas complet empire le score
        scale, q_try = 1.0, None
        for _ in range(3):
            q_try = clamp([q[j] + scale * dq[j] for j in range(6)])
            Pt = fk_pose(q_try)
            ept = [tpos[i] - eff_pos(Pt)[i] for i in range(3)]
            eot = ori_err(cols(Pt), RG)
            st = math.sqrt(sum(v*v for v in ept)) + wo * math.sqrt(sum(v*v for v in eot))
            if st < s:
                break
            scale *= 0.5
        q = q_try
    P = fk_pose(best_q)
    rp = math.sqrt(sum((tpos[i] - eff_pos(P)[i])**2 for i in range(3)))
    ro = math.degrees(math.sqrt(sum(v*v for v in ori_err(cols(P), RG))))
    return best_q, rp, ro


def applique(q):
    for (nom, axe, lo, hi), a in zip(ARM, q):
        F[nom].setPose(REST[nom] * ROT[axe](math.radians(a)))


# ---------------- choregraphie v3 : cles -> trajectoire precalculee ------
cube_y = TABLE_TOP + CUBE / 2.0          # centre du cube
GRASP_Y = cube_y + CUBE / 2.0 + GRASP_CLEAR   # centre main, cube en main

q_rest = [0.0] * 6

# Cles FK de la MONTEE : le coude PART EN ARRIERE (flexion epaule
# positive) pendant que le pli du coude monte la main devant la poitrine.
# L'epaule part FRANCHEMENT en extension (+34/+36) des l'amorce : pendant
# le pli, l'arc de l'avant-bras balaie vers l'avant, et la face avant de
# la table n'est qu'a 50 mm de la main au repos — epaule a +14 ca frotte
# (17 collisions mesh), a +34 ca passe (0, banc _tune_keys). La descente
# du retour reutilise ces cles en miroir.
QK_A = [-6.0, 34.0, 5.0, -30.0, -30.0, 0.0]    # amorce : epaule bien ARRIERE
QK_B = [-12.0, 36.0, 10.0, -95.0, -35.0, 0.0]  # main haute pres du corps

# Cibles cartesiennes (resolues en cles articulaires par IK, HORS animation)
P_PREPICK = (PICK_X, GRASP_Y + 35, PICK_Z - 10)
P_PICK = (PICK_X, GRASP_Y, PICK_Z)
P_HI_PICK = (PICK_X, HI, TRANSIT_Z)
P_HI_MID = ((PICK_X + PLACE_X) / 2.0, HI, TRANSIT_Z)
P_HI_PLACE = (PLACE_X, HI, TRANSIT_Z)
P_PLACE = (PLACE_X, GRASP_Y, PLACE_Z)

# phases : (label, vitesse deg/frame, pause_s, evenement_de_fin)
# Les cles de chaque phase sont resolues dans build_trajectoire().
# Le rendu RoboDK coute ~80 ms/frame (mesure 11/06) : c'est LUI la cadence
# reelle, pas DT. Les pas sont donc dimensionnes pour un geste dynamique a
# ~12 fps rendus : 6 deg/frame ~ 70 deg/s effectifs sur les grands gestes.
V_VIF = 6.0      # deg max/frame pour les grands gestes
V_FIN = 3.0      # approche / depose : plus pose


def _dist(a, b):
    return math.sqrt(sum((x - y) ** 2 for x, y in zip(a, b)))


def catmull(pts, u):
    """Point sur la spline Catmull-Rom 6D passant par pts (u dans [0,1],
    parametrisation par longueur de corde). 2 points = segment droit."""
    P = [pts[0]] + list(pts) + [pts[-1]]
    L = [_dist(pts[i], pts[i + 1]) for i in range(len(pts) - 1)]
    tot = sum(L) or 1.0
    s = u * tot
    i = 0
    while i < len(L) - 1 and s > L[i]:
        s -= L[i]
        i += 1
    t = s / (L[i] or 1.0)
    p0, p1, p2, p3 = P[i], P[i + 1], P[i + 2], P[i + 3]
    return [0.5 * (2 * p1[k] + (-p0[k] + p2[k]) * t
                   + (2 * p0[k] - 5 * p1[k] + 4 * p2[k] - p3[k]) * t * t
                   + (-p0[k] + 3 * p1[k] - 3 * p2[k] + p3[k]) * t ** 3)
            for k in range(len(pts[0]))]


def _resample(keys, v_frame):
    """Echantillonne la spline articulaire passant par keys en frames a
    vitesse bornee : nombre de frames dimensionne sur le plus grand ecart
    articulaire, profil smoothstep (doux au depart et a l'arrivee)."""
    span = 0.0
    for a, b in zip(keys, keys[1:]):
        span += max(abs(x - y) for x, y in zip(a, b))
    n = max(4, int(math.ceil(span / v_frame)))
    out = []
    for s in range(1, n + 1):
        t = s / n
        t = t * t * (3 - 2 * t)                  # smoothstep
        out.append(clamp(catmull(keys, t)))
    return out


def build_trajectoire():
    """Resout toutes les cles (IK hors animation) puis precalcule TOUTES
    les frames. Retourne (frames, events, rapport) avec
    frames = [q, ...], events = {index_frame: nom}, et un rapport texte
    (residus IK + scan coude)."""
    rapport = []

    def cle_ik(nom, cible, q_seed, wo):
        q, rp, ro = ik(cible, q_seed, wo=wo)
        rapport.append(f"  cle {nom:<10} residu {rp:5.1f} mm / {ro:5.1f} deg")
        if rp > 14:
            rapport.append(f"    !! {nom} : cible mal atteinte ({rp:.0f} mm)")
        return q

    # pick d'abord (seed = cle FK de la montee), puis prepick ANCRE sur la
    # branche de pick (meme poids d'orientation) : sans ca, l'approche
    # lente traversait un saut de branche (poignet -16 -> +50 deg).
    q_pick = cle_ik("pick", P_PICK, QK_B, WO)
    q_prepick = cle_ik("prepick", P_PREPICK, q_pick, WO)
    q_hi1 = cle_ik("hi_pick", P_HI_PICK, q_pick, WO)
    q_him = cle_ik("hi_mid", P_HI_MID, q_hi1, WO)
    q_hi2 = cle_ik("hi_place", P_HI_PLACE, q_him, WO)
    q_place = cle_ik("place", P_PLACE, q_hi2, WO)

    phases = [
        ("tendre", [q_rest, QK_A, QK_B, q_prepick], V_VIF, 0.0, None),
        ("saisir", [q_prepick, q_pick], V_FIN, 0.30, "grab"),
        ("transporter", [q_pick, q_hi1, q_him, q_hi2], V_VIF, 0.0, None),
        ("deposer", [q_hi2, q_place], V_FIN, 0.30, "release"),
        ("ramener", [q_place, q_hi2, QK_B, QK_A, q_rest], V_VIF, 0.0, None),
    ]

    frames, events, pauses = [], {}, {}
    for label, keys, v, pause, event in phases:
        fr = _resample(keys, v)
        frames += fr
        if event:
            events[len(frames) - 1] = event
        if pause:
            pauses[len(frames) - 1] = pause
        rapport.append(f"  phase {label:<12} {len(fr):3d} frames")

    # SCAN COUDE : garantie "jamais en avant" sur la trajectoire COMPLETE
    z0 = fk_coude(q_rest)[2]
    zmax, imax = -1e9, 0
    for i, q in enumerate(frames):
        z = fk_coude(q)[2]
        if z > zmax:
            zmax, imax = z, i
    ok = zmax <= z0 + 5.0
    rapport.append(f"  coude : Z repos {z0:.0f} mm, Z max trajectoire "
                   f"{zmax:.0f} mm (frame {imax}) -> "
                   f"{'OK, jamais en avant' if ok else '!! PART EN AVANT'}")
    return frames, events, pauses, rapport, ok


def main():
    print("--- Tache bras v3 : coude en arriere, trajectoire precalculee ---")
    t0 = time.time()
    frames, events, pauses, rapport, coude_ok = build_trajectoire()
    print("\n".join(rapport))
    print(f"Precalcul : {len(frames)} frames en {time.time() - t0:.1f} s "
          f"(~{len(frames) * DT + sum(pauses.values()):.1f} s d'animation)")
    if not coude_ok:
        sys.exit("ABANDON : le coude partirait en avant — cles a corriger.")
    if "--check" in sys.argv:
        print("--check : pas d'animation.")
        return

    station = RDK.ActiveStation()
    wrist = F[ARM[-1][0]]
    if "--frames" not in sys.argv:            # demo propre : cacher les reperes
        for fr in RDK.ItemList(ITEM_TYPE_FRAME):
            fr.setVisible(False, False)
    piece.setParentStatic(station)            # remettre la piece au depart
    piece.setPose(transl(PICK_X, cube_y, PICK_Z))
    applique(q_rest)
    RDK.Render(True)
    time.sleep(0.3)

    # LECTURE : zero calcul, cadence reelle tenue sur l'horloge murale
    # (si le rendu prend du retard, on saute le sleep, pas des frames).
    t0 = time.time()
    for i, q in enumerate(frames):
        applique(q)
        RDK.Render(True)
        ev = events.get(i)
        if ev == "grab":
            piece.setParentStatic(wrist)      # la piece suit la main
            print("  piece saisie")
        elif ev == "release":
            piece.setParentStatic(station)
            piece.setPose(transl(PLACE_X, cube_y, PLACE_Z))
            print(f"  piece deposee en ({PLACE_X:.0f}, {cube_y:.0f}, {PLACE_Z:.0f})")
        if i in pauses:
            time.sleep(pauses[i])
            t0 += pauses[i]
        reste = t0 + (i + 1) * DT - time.time()
        if reste > 0:
            time.sleep(reste)
    print(f"Fini en {time.time() - t0:.1f} s - piece deplacee de gauche a "
          f"droite, coude toujours en arriere.")


if __name__ == "__main__":
    main()
